// TIA Portal V21 export
// export: Created 2026-10-27T23:04:39.0346325Z, ExportSetting WithDefaults, DisplayName Totally Integrated Automation Portal, DisplayVersion V21 Update 3, DisplayName TIA Portal Test Suite Advanced, DisplayVersion V21 Update 1, DisplayName SINAMICS Startdrive Advanced, DisplayVersion V21 Update 1, DisplayName SINAMICS Startdrive G130, G150, S120, S150, G200, G210, G210C, G210X, G220, S200, S210, S220, Innomotics MVD, DisplayVersion V21 Update 1, DisplayName SINAMICS Startdrive G110M, G120, G120C, G120D, G120P, G115D, DisplayVersion V21 Update 1, DisplayName STEP 7 Professional, DisplayVersion V21 Update 3, DisplayName STEP 7 Safety, DisplayVersion V21, DisplayName Tech WebApplication, DisplayVersion V21, DisplayName WinCC Basic/Comfort/Advanced, DisplayVersion V21 Update 3, DisplayName WinCC Professional, DisplayVersion V21 Update 3, DisplayName WinCC Unified, DisplayVersion V21 Update 3
FUNCTION_BLOCK "Tgp_MulReal_FBD"   // FB29, FBD
{ S7_Optimized_Access := 'TRUE' }
VERSION : 0.1
// stored: AutoNumber true, IsIECCheckEnabled false, IsRetainMemResEnabled false, MemoryReserve 100, SetENOAutomatically false, UDAEnableTagReadback false
   VAR_INPUT
      Left : Real;
      Right : Real;
   END_VAR
   VAR_OUTPUT
      Result : Real;
   END_VAR
BEGIN

REGION Network 1
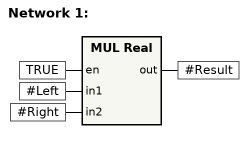
   IF TRUE THEN #Result := #Left * #Right; END_IF;
END_REGION
END_FUNCTION_BLOCK
